(* Logix 5000 project; controller R400_500_XLS vendor 1 type 14 code 216 rev 31.11; software revision 31.01; part 15 of 32 *)
(* tags used below, declared in another part *)
   CycleModifBuffer : UDT_CYCLE;
   CycleNotEmpty : SINT;
   First_Inj_conc : BOOL;
   M : DINT[5];   // Memory Bits
   MaxTrtTempSp : REAL;
   PreWash_Select : BOOL;
   PrewashIndex : SINT;   // Index of the selected pre-wash treatment
   Rinse_Select : BOOL;
   RinseIndex : SINT;
   Second_Inj_conc : BOOL;
   Tmr : TIMER[107];
   Wash_Select : BOOL;
   WashIndex : SINT;
   WashInjectionType1 : DINT;
   CfgChem : SINT;
   CfgChem2 : SINT;
   CfgConc : REAL;
   CfgConc2 : REAL;
   CfgCondSp : REAL;
   CfgInjType : SINT;
   cfgPrewashHeated : SINT;
   cfgPrewashMin : SINT;
   cfgPrewashSec : DINT;
   CfgPrewashTempSp : REAL;
   CfgWshHeated : SINT;
   CfgWshInjRateImperial : REAL;   // Wash Injection Rate - Oz / Gal
   CfgWshInjRateMetric : REAL;   // Wash Injection Rate - mL / L
   CfgWshMin : SINT;
   CfgWshSec : SINT;
   CfgWshTempSp : REAL;
   cfgWshWport : SINT;
   ChemConcUnit : BOOL;   // 0 = mL/L; 1 = oz/gal
   Msg_TempSp : SINT;   // HMI Information Message tag
   Msg_TempSp_Ack : BOOL;
   NumInput : UDT_NUMERIC_INPUT[65];   // Numeric input
   NumInputReal : UDT_NUMERIC_INPUT_REAL[17];
   Screen_Ctrl : DINT;   // PLC Screen Request
   Selector : UDT_SELECTOR[25];   // Piloted list selector
   TempUnit : BOOL;   // Temperature Units 0= Celcius 1 = Farhenheit
   Tpb : DINT[11];
   TpbImage : DINT[11];
(* MainProgram, continued *)

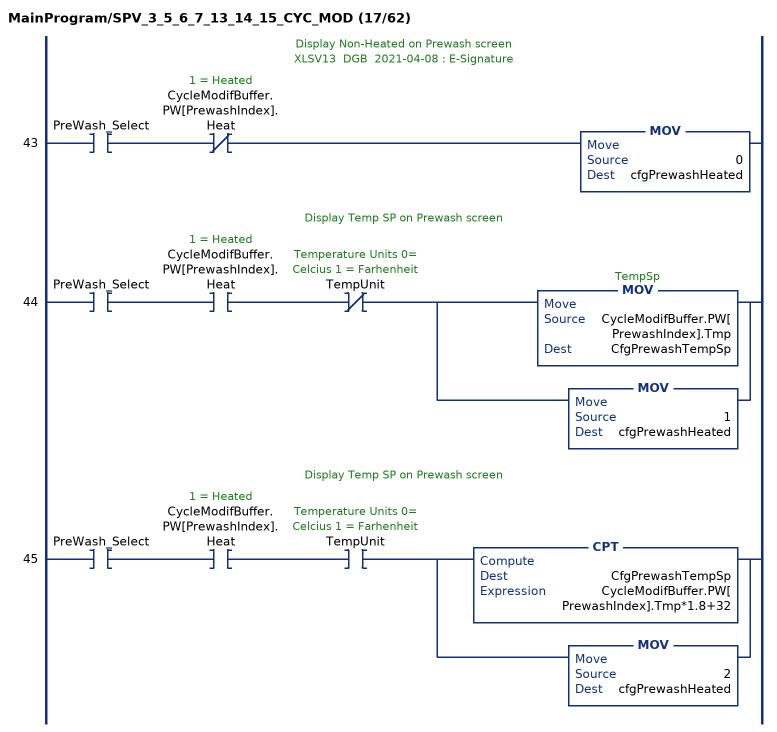
   [picture p268: MainProgram/SPV_3_5_6_7_13_14_15_CYC_MOD rungs 43-45]
   // Display Non-Heated on Prewash screen
   // XLSV13  DGB  2021-04-08 : E-Signature
   43: XIC(PreWash_Select)XIO(CycleModifBuffer.PW[PrewashIndex].Heat)MOV(0,cfgPrewashHeated);
   // Display Temp SP on Prewash screen
   44: XIC(PreWash_Select)XIC(CycleModifBuffer.PW[PrewashIndex].Heat)XIO(TempUnit)[MOV(CycleModifBuffer.PW[PrewashIndex].Tmp,CfgPrewashTempSp) ,MOV(1,cfgPrewashHeated) ];
   // Display Temp SP on Prewash screen
   45: XIC(PreWash_Select)XIC(CycleModifBuffer.PW[PrewashIndex].Heat)XIC(TempUnit)[CPT(CfgPrewashTempSp,CycleModifBuffer.PW[PrewashIndex].Tmp*1.8+32) ,MOV(2,cfgPrewashHeated) ];
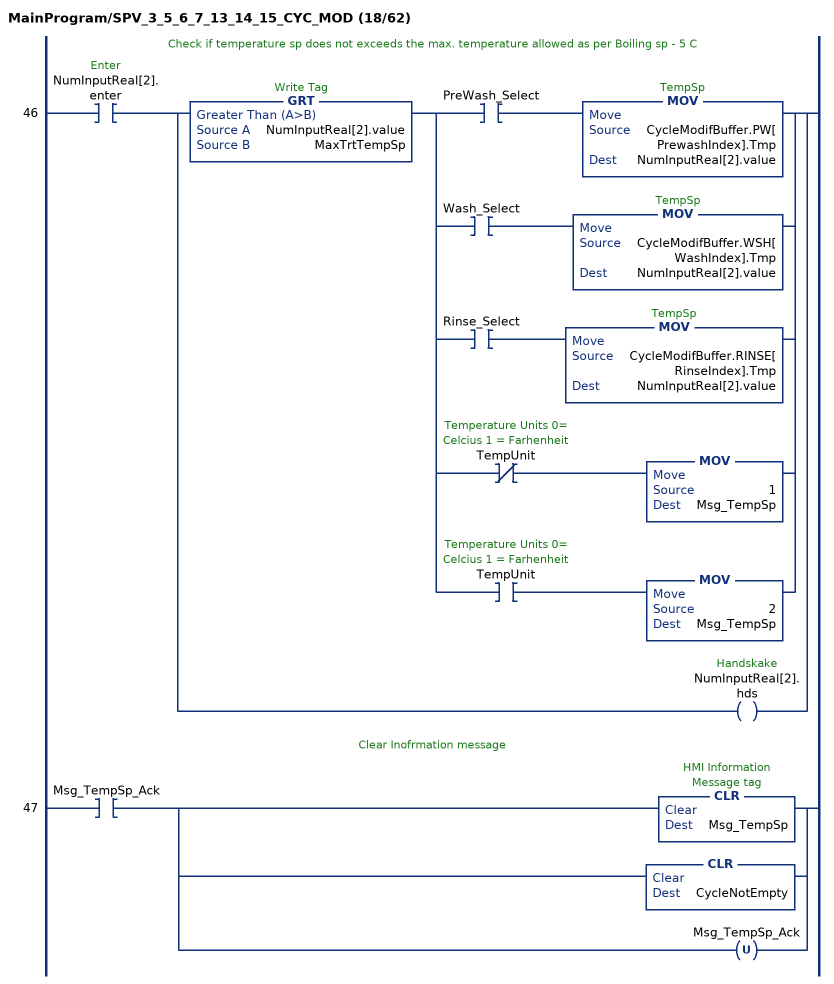
   // Check if temperature sp does not exceeds the max. temperature allowed as per Boiling sp - 5 C
   46: XIC(NumInputReal[2].enter)[GRT(NumInputReal[2].value,MaxTrtTempSp) [XIC(PreWash_Select) MOV(CycleModifBuffer.PW[PrewashIndex].Tmp,NumInputReal[2].value) ,XIC(Wash_Select) MOV(CycleModifBuffer.WSH[WashIndex].Tmp,NumInputReal[2].value) ,XIC(Rinse_Select) MOV(CycleModifBuffer.RINSE[RinseIndex].Tmp,NumInputReal[2].value) ,XIO(TempUnit) MOV(1,Msg_TempSp) ,XIC(TempUnit) MOV(2,Msg_TempSp) ] ,OTE(NumInputReal[2].hds) ];
   // Clear Inofrmation message
   47: XIC(Msg_TempSp_Ack)[CLR(Msg_TempSp) ,CLR(CycleNotEmpty) ,OTU(Msg_TempSp_Ack) ];
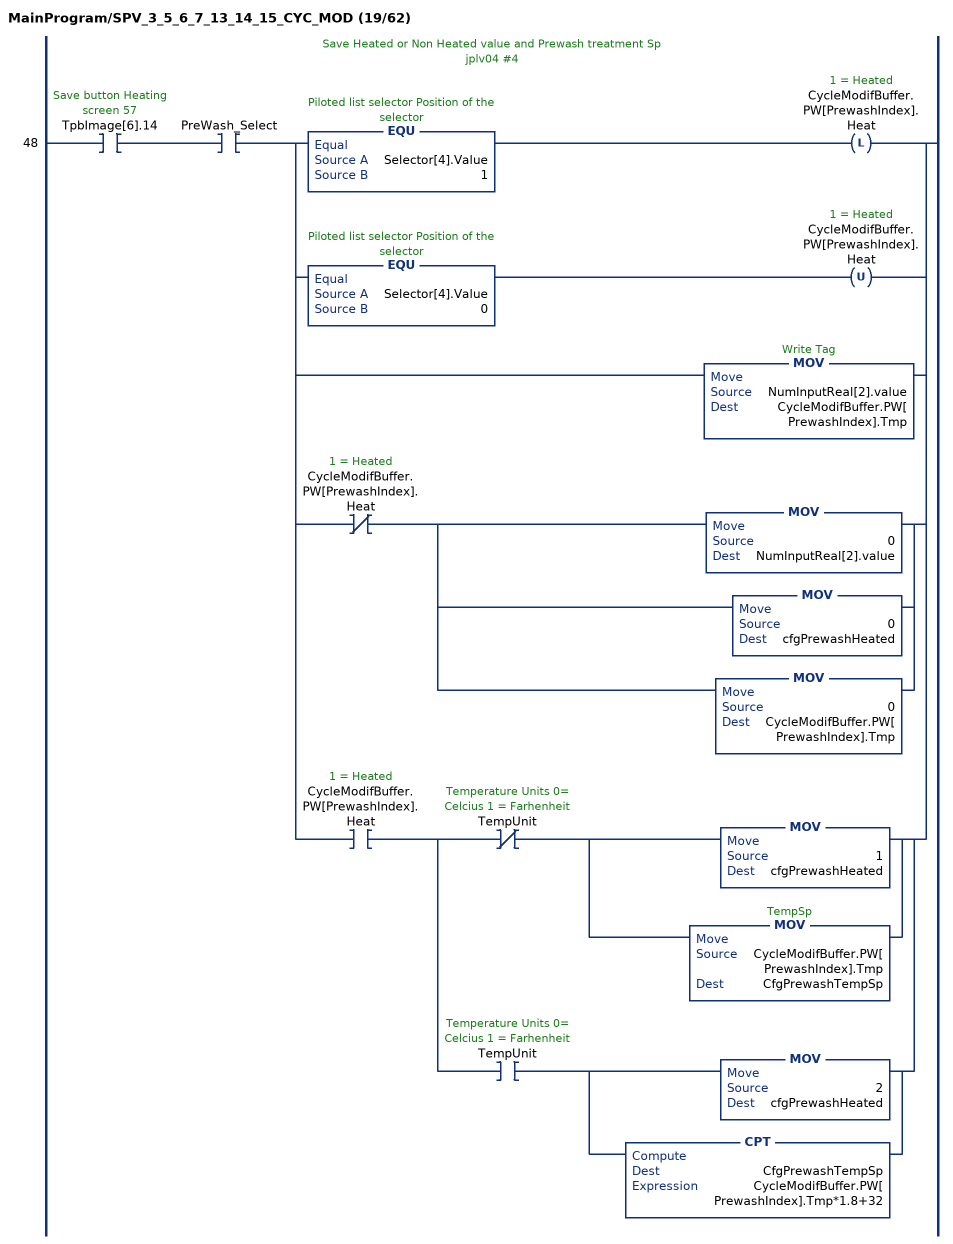
   // Save Heated or Non Heated value and Prewash treatment Sp
   // jplv04 #4
   48: XIC(TpbImage[6].14)XIC(PreWash_Select)[EQU(Selector[4].Value,1) OTL(CycleModifBuffer.PW[PrewashIndex].Heat) ,EQU(Selector[4].Value,0) OTU(CycleModifBuffer.PW[PrewashIndex].Heat) ,MOV(NumInputReal[2].value,CycleModifBuffer.PW[PrewashIndex].Tmp) ,XIO(CycleModifBuffer.PW[PrewashIndex].Heat) [MOV(0,NumInputReal[2].value) ,MOV(0,cfgPrewashHeated) ,MOV(0,CycleModifBuffer.PW[PrewashIndex].Tmp) ] ,XIC(CycleModifBuffer.PW[PrewashIndex].Heat) [XIO(TempUnit) [MOV(1,cfgPrewashHeated) ,MOV(CycleModifBuffer.PW[PrewashIndex].Tmp,CfgPrewashTempSp) ] ,XIC(TempUnit) [MOV(2,cfgPrewashHeated) ,CPT(CfgPrewashTempSp,CycleModifBuffer.PW[PrewashIndex].Tmp*1.8+32) ] ] ];
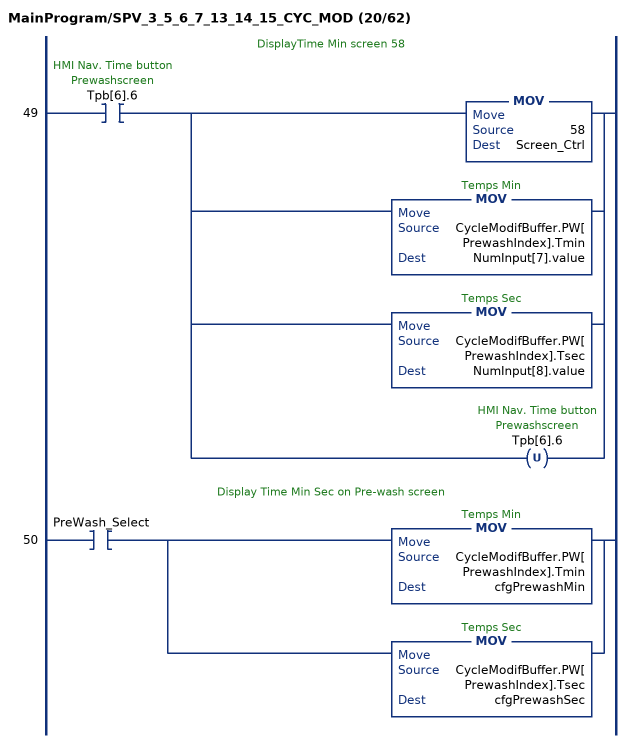
   // DisplayTime Min screen 58
   49: XIC(Tpb[6].6)[MOV(58,Screen_Ctrl) ,MOV(CycleModifBuffer.PW[PrewashIndex].Tmin,NumInput[7].value) ,MOV(CycleModifBuffer.PW[PrewashIndex].Tsec,NumInput[8].value) ,OTU(Tpb[6].6) ];
   // Display Time Min Sec on Pre-wash screen
   50: XIC(PreWash_Select)[MOV(CycleModifBuffer.PW[PrewashIndex].Tmin,cfgPrewashMin) ,MOV(CycleModifBuffer.PW[PrewashIndex].Tsec,cfgPrewashSec) ];
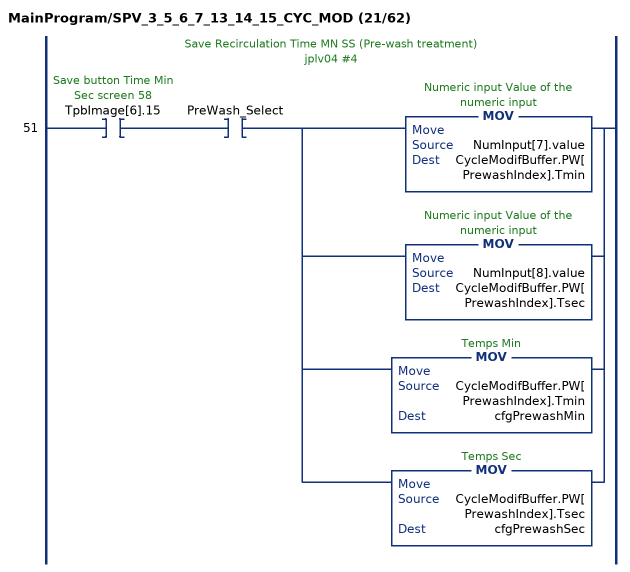
   // Save Recirculation Time MN SS (Pre-wash treatment)
   // jplv04 #4
   51: XIC(TpbImage[6].15)XIC(PreWash_Select)[MOV(NumInput[7].value,CycleModifBuffer.PW[PrewashIndex].Tmin) ,MOV(NumInput[8].value,CycleModifBuffer.PW[PrewashIndex].Tsec) ,MOV(CycleModifBuffer.PW[PrewashIndex].Tmin,cfgPrewashMin) ,MOV(CycleModifBuffer.PW[PrewashIndex].Tsec,cfgPrewashSec) ];
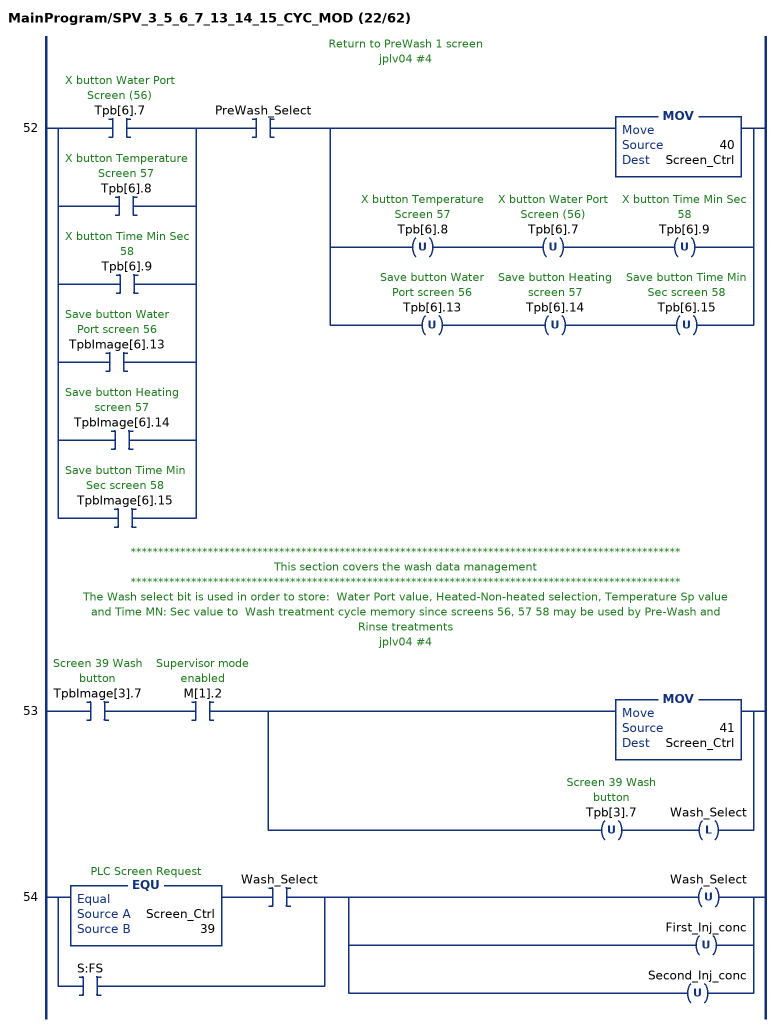
   // Return to PreWash 1 screen
   // jplv04 #4
   52: [XIC(Tpb[6].7) ,XIC(Tpb[6].8) ,XIC(Tpb[6].9) ,XIC(TpbImage[6].13) ,XIC(TpbImage[6].14) ,XIC(TpbImage[6].15) ]XIC(PreWash_Select)[MOV(40,Screen_Ctrl) ,OTU(Tpb[6].8) OTU(Tpb[6].7) OTU(Tpb[6].9) ,OTU(Tpb[6].13) OTU(Tpb[6].14) OTU(Tpb[6].15) ];
   // ****************************************************************************************************
   // This section covers the wash data management
   // ****************************************************************************************************
   // The Wash select bit is used in order to store:  Water Port value, Heated-Non-heated selection, Temperature Sp value and Time MN: Sec value to  Wash treatment cycle memory since screens 56, 57 58 may be used by Pre-Wash and Rinse treatments
   // jplv04 #4
   53: XIC(TpbImage[3].7)XIC(M[1].2)[MOV(41,Screen_Ctrl) ,OTU(Tpb[3].7) OTL(Wash_Select) ];
   54: [EQU(Screen_Ctrl,39) XIC(Wash_Select) ,XIC(S:FS) ][OTU(Wash_Select) ,OTU(First_Inj_conc) ,OTU(Second_Inj_conc) ];
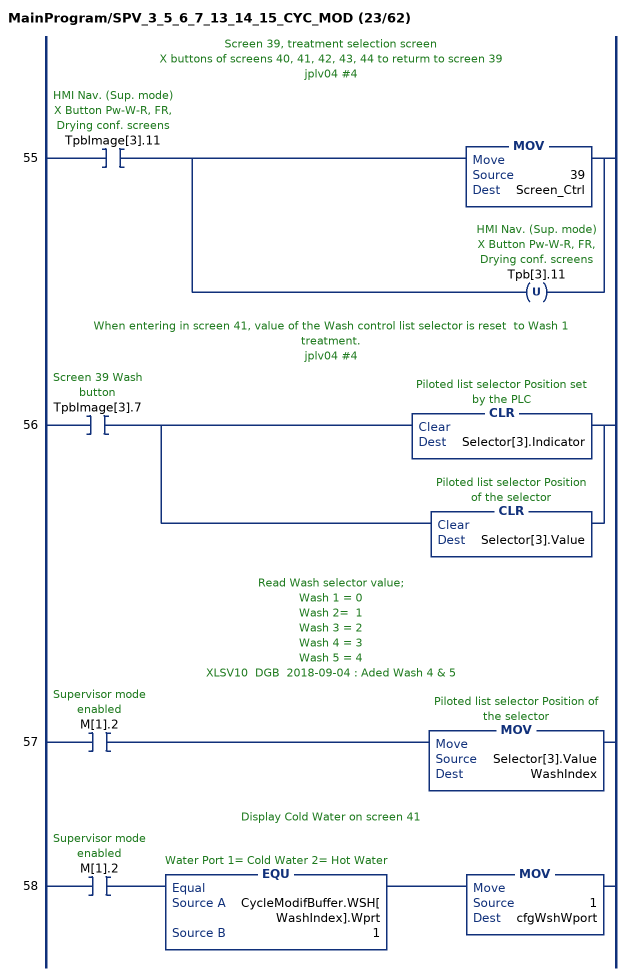
   // Screen 39, treatment selection screen
   // X buttons of screens 40, 41, 42, 43, 44 to returm to screen 39
   // jplv04 #4
   55: XIC(TpbImage[3].11)[MOV(39,Screen_Ctrl) ,OTU(Tpb[3].11) ];
   // When entering in screen 41, value of the Wash control list selector is reset  to Wash 1 treatment.
   // jplv04 #4
   56: XIC(TpbImage[3].7)[CLR(Selector[3].Indicator) ,CLR(Selector[3].Value) ];
   // Read Wash selector value;
   // Wash 1 = 0
   // Wash 2=  1
   // Wash 3 = 2
   // Wash 4 = 3
   // Wash 5 = 4
   // XLSV10  DGB  2018-09-04 : Aded Wash 4 & 5
   57: XIC(M[1].2)MOV(Selector[3].Value,WashIndex);
   // Display Cold Water on screen 41
   58: XIC(M[1].2)EQU(CycleModifBuffer.WSH[WashIndex].Wprt,1)MOV(1,cfgWshWport);
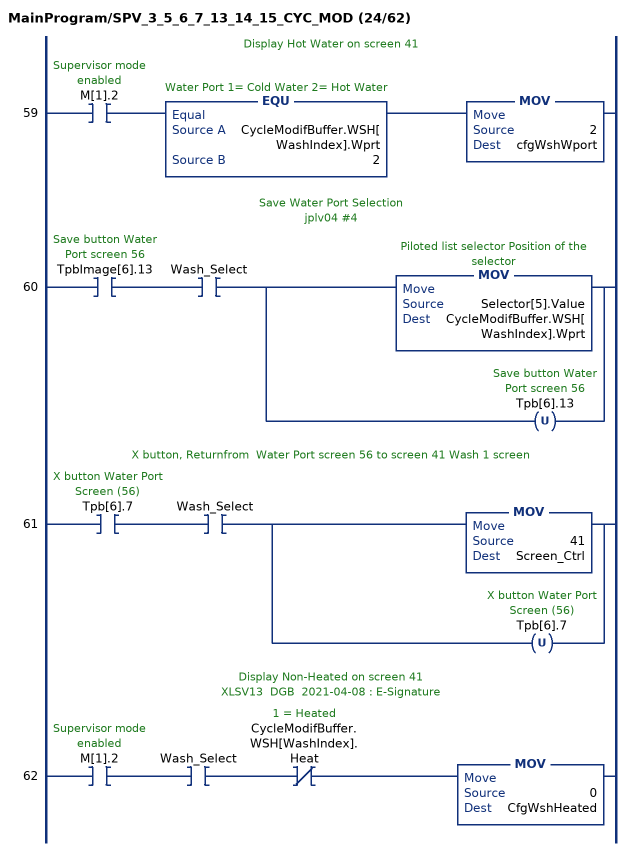
   // Display Hot Water on screen 41
   59: XIC(M[1].2)EQU(CycleModifBuffer.WSH[WashIndex].Wprt,2)MOV(2,cfgWshWport);
   // Save Water Port Selection
   // jplv04 #4
   60: XIC(TpbImage[6].13)XIC(Wash_Select)[MOV(Selector[5].Value,CycleModifBuffer.WSH[WashIndex].Wprt) ,OTU(Tpb[6].13) ];
   // X button, Returnfrom  Water Port screen 56 to screen 41 Wash 1 screen
   61: XIC(Tpb[6].7)XIC(Wash_Select)[MOV(41,Screen_Ctrl) ,OTU(Tpb[6].7) ];
   // Display Non-Heated on screen 41
   // XLSV13  DGB  2021-04-08 : E-Signature
   62: XIC(M[1].2)XIC(Wash_Select)XIO(CycleModifBuffer.WSH[WashIndex].Heat)MOV(0,CfgWshHeated);
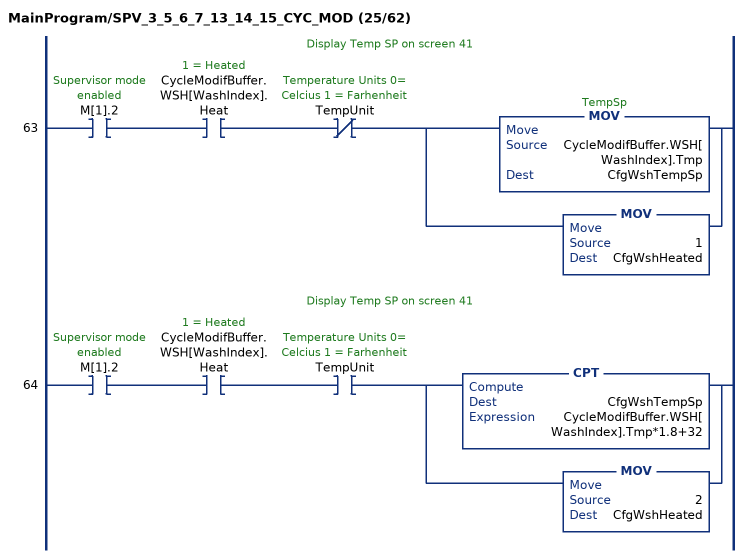
   // Display Temp SP on screen 41
   63: XIC(M[1].2)XIC(CycleModifBuffer.WSH[WashIndex].Heat)XIO(TempUnit)[MOV(CycleModifBuffer.WSH[WashIndex].Tmp,CfgWshTempSp) ,MOV(1,CfgWshHeated) ];
   // Display Temp SP on screen 41
   64: XIC(M[1].2)XIC(CycleModifBuffer.WSH[WashIndex].Heat)XIC(TempUnit)[CPT(CfgWshTempSp,CycleModifBuffer.WSH[WashIndex].Tmp*1.8+32) ,MOV(2,CfgWshHeated) ];
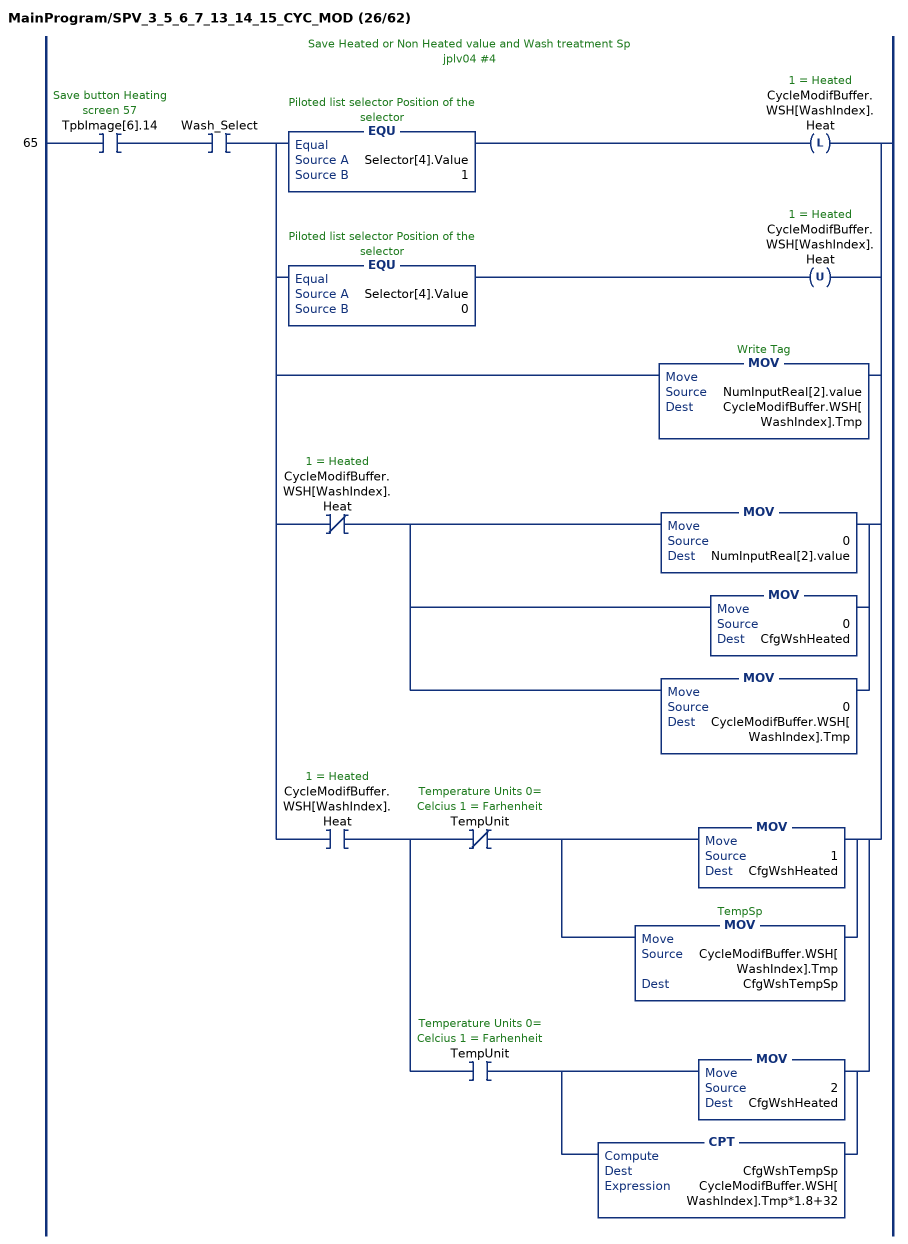
   // Save Heated or Non Heated value and Wash treatment Sp
   // jplv04 #4
   65: XIC(TpbImage[6].14)XIC(Wash_Select)[EQU(Selector[4].Value,1) OTL(CycleModifBuffer.WSH[WashIndex].Heat) ,EQU(Selector[4].Value,0) OTU(CycleModifBuffer.WSH[WashIndex].Heat) ,MOV(NumInputReal[2].value,CycleModifBuffer.WSH[WashIndex].Tmp) ,XIO(CycleModifBuffer.WSH[WashIndex].Heat) [MOV(0,NumInputReal[2].value) ,MOV(0,CfgWshHeated) ,MOV(0,CycleModifBuffer.WSH[WashIndex].Tmp) ] ,XIC(CycleModifBuffer.WSH[WashIndex].Heat) [XIO(TempUnit) [MOV(1,CfgWshHeated) ,MOV(CycleModifBuffer.WSH[WashIndex].Tmp,CfgWshTempSp) ] ,XIC(TempUnit) [MOV(2,CfgWshHeated) ,CPT(CfgWshTempSp,CycleModifBuffer.WSH[WashIndex].Tmp*1.8+32) ] ] ];
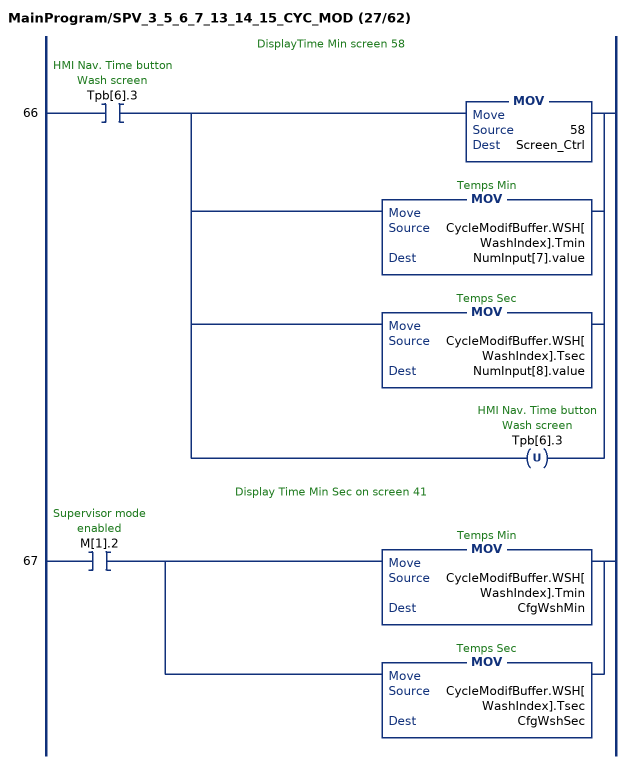
   // DisplayTime Min screen 58
   66: XIC(Tpb[6].3)[MOV(58,Screen_Ctrl) ,MOV(CycleModifBuffer.WSH[WashIndex].Tmin,NumInput[7].value) ,MOV(CycleModifBuffer.WSH[WashIndex].Tsec,NumInput[8].value) ,OTU(Tpb[6].3) ];
   // Display Time Min Sec on screen 41
   67: XIC(M[1].2)[MOV(CycleModifBuffer.WSH[WashIndex].Tmin,CfgWshMin) ,MOV(CycleModifBuffer.WSH[WashIndex].Tsec,CfgWshSec) ];
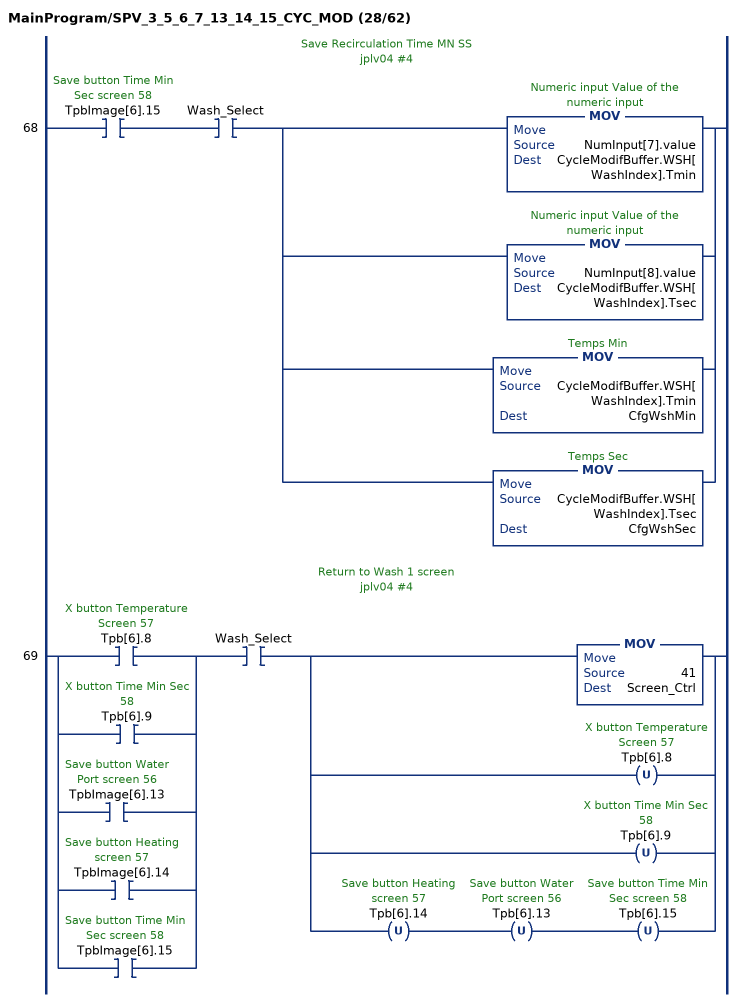
   // Save Recirculation Time MN SS
   // jplv04 #4
   68: XIC(TpbImage[6].15)XIC(Wash_Select)[MOV(NumInput[7].value,CycleModifBuffer.WSH[WashIndex].Tmin) ,MOV(NumInput[8].value,CycleModifBuffer.WSH[WashIndex].Tsec) ,MOV(CycleModifBuffer.WSH[WashIndex].Tmin,CfgWshMin) ,MOV(CycleModifBuffer.WSH[WashIndex].Tsec,CfgWshSec) ];
   // Return to Wash 1 screen
   // jplv04 #4
   69: [XIC(Tpb[6].8) ,XIC(Tpb[6].9) ,XIC(TpbImage[6].13) ,XIC(TpbImage[6].14) ,XIC(TpbImage[6].15) ]XIC(Wash_Select)[MOV(41,Screen_Ctrl) ,OTU(Tpb[6].8) ,OTU(Tpb[6].9) ,OTU(Tpb[6].14) OTU(Tpb[6].13) OTU(Tpb[6].15) ];
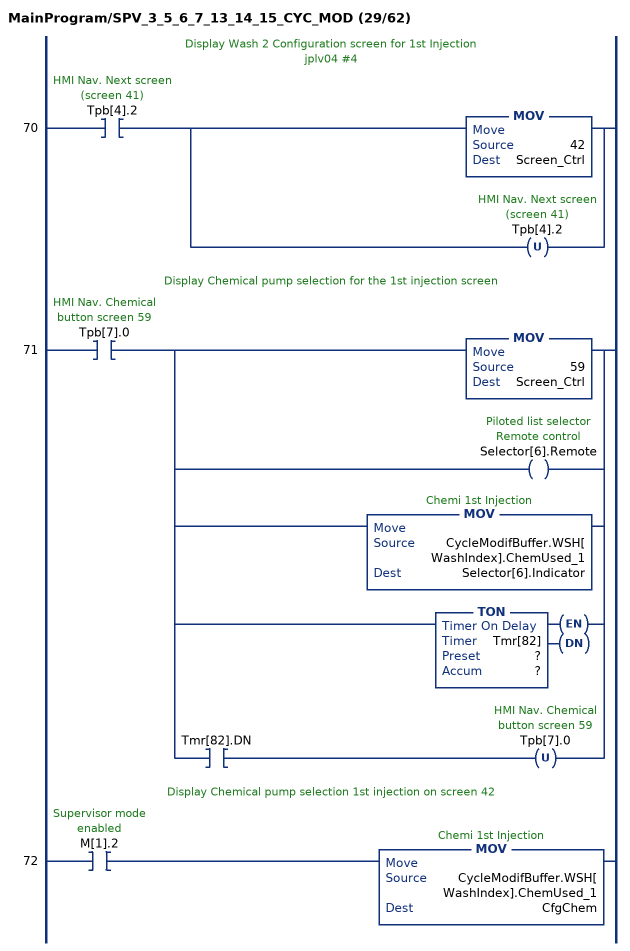
   // Display Wash 2 Configuration screen for 1st Injection
   // jplv04 #4
   70: XIC(Tpb[4].2)[MOV(42,Screen_Ctrl) ,OTU(Tpb[4].2) ];
   // Display Chemical pump selection for the 1st injection screen
   71: XIC(Tpb[7].0)[MOV(59,Screen_Ctrl) ,OTE(Selector[6].Remote) ,MOV(CycleModifBuffer.WSH[WashIndex].ChemUsed_1,Selector[6].Indicator) ,TON(Tmr[82],?,?) ,XIC(Tmr[82].DN) OTU(Tpb[7].0) ];
   // Display Chemical pump selection 1st injection on screen 42
   72: XIC(M[1].2)MOV(CycleModifBuffer.WSH[WashIndex].ChemUsed_1,CfgChem);
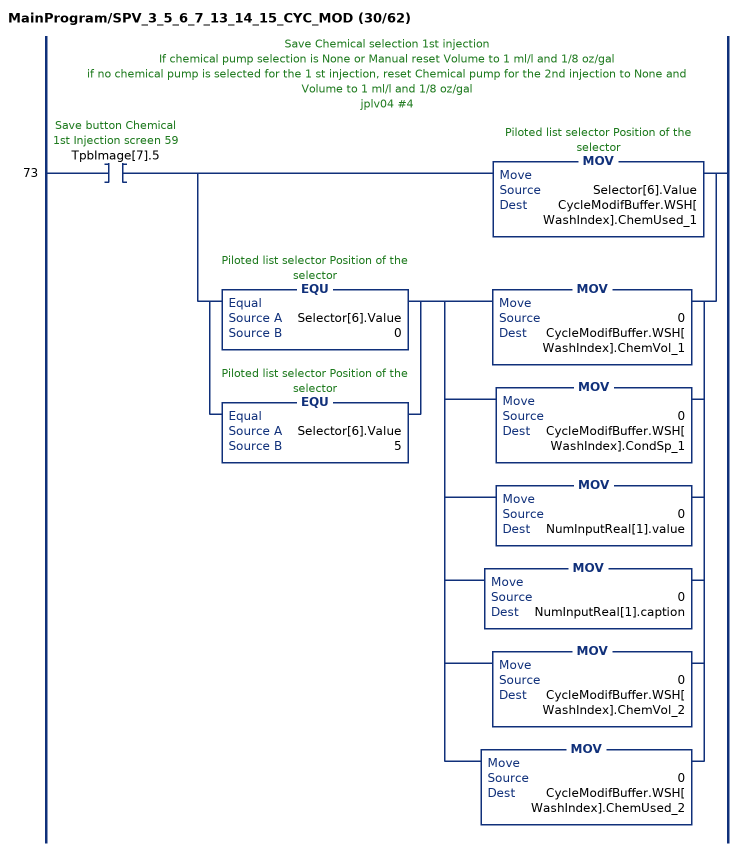
   // Save Chemical selection 1st injection
   // If chemical pump selection is None or Manual reset Volume to 1 ml/l and 1/8 oz/gal
   // if no chemical pump is selected for the 1 st injection, reset Chemical pump for the 2nd injection to None and Volume to 1 ml/l and 1/8 oz/gal
   // jplv04 #4
   73: XIC(TpbImage[7].5)[MOV(Selector[6].Value,CycleModifBuffer.WSH[WashIndex].ChemUsed_1) ,[EQU(Selector[6].Value,0) ,EQU(Selector[6].Value,5) ] [MOV(0,CycleModifBuffer.WSH[WashIndex].ChemVol_1) ,MOV(0,CycleModifBuffer.WSH[WashIndex].CondSp_1) ,MOV(0,NumInputReal[1].value) ,MOV(0,NumInputReal[1].caption) ,MOV(0,CycleModifBuffer.WSH[WashIndex].ChemVol_2) ,MOV(0,CycleModifBuffer.WSH[WashIndex].ChemUsed_2) ] ];
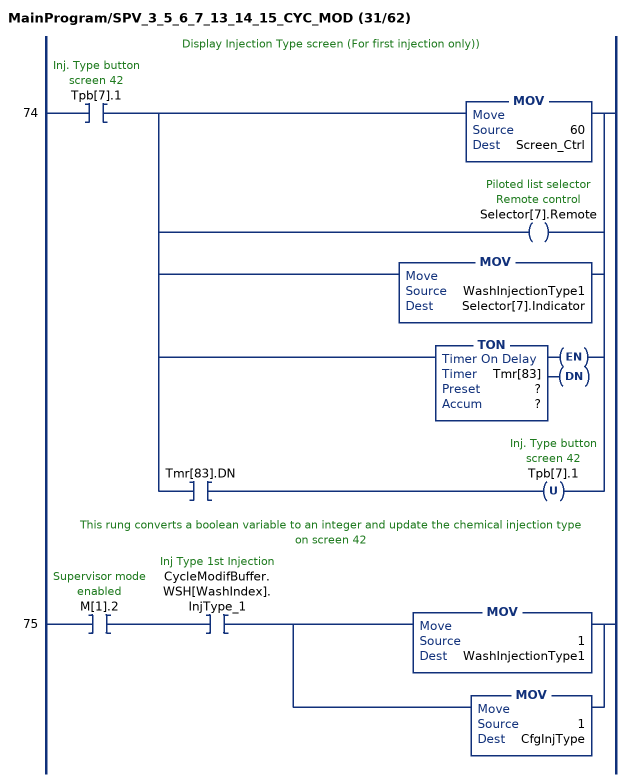
   // Display Injection Type screen (For first injection only))
   74: XIC(Tpb[7].1)[MOV(60,Screen_Ctrl) ,OTE(Selector[7].Remote) ,MOV(WashInjectionType1,Selector[7].Indicator) ,TON(Tmr[83],?,?) ,XIC(Tmr[83].DN) OTU(Tpb[7].1) ];
   // This rung converts a boolean variable to an integer and update the chemical injection type on screen 42
   75: XIC(M[1].2)XIC(CycleModifBuffer.WSH[WashIndex].InjType_1)[MOV(1,WashInjectionType1) ,MOV(1,CfgInjType) ];
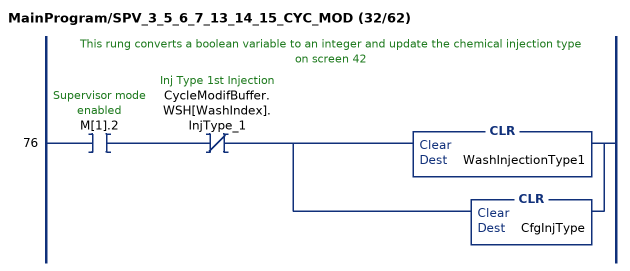
   // This rung converts a boolean variable to an integer and update the chemical injection type on screen 42
   76: XIC(M[1].2)XIO(CycleModifBuffer.WSH[WashIndex].InjType_1)[CLR(WashInjectionType1) ,CLR(CfgInjType) ];
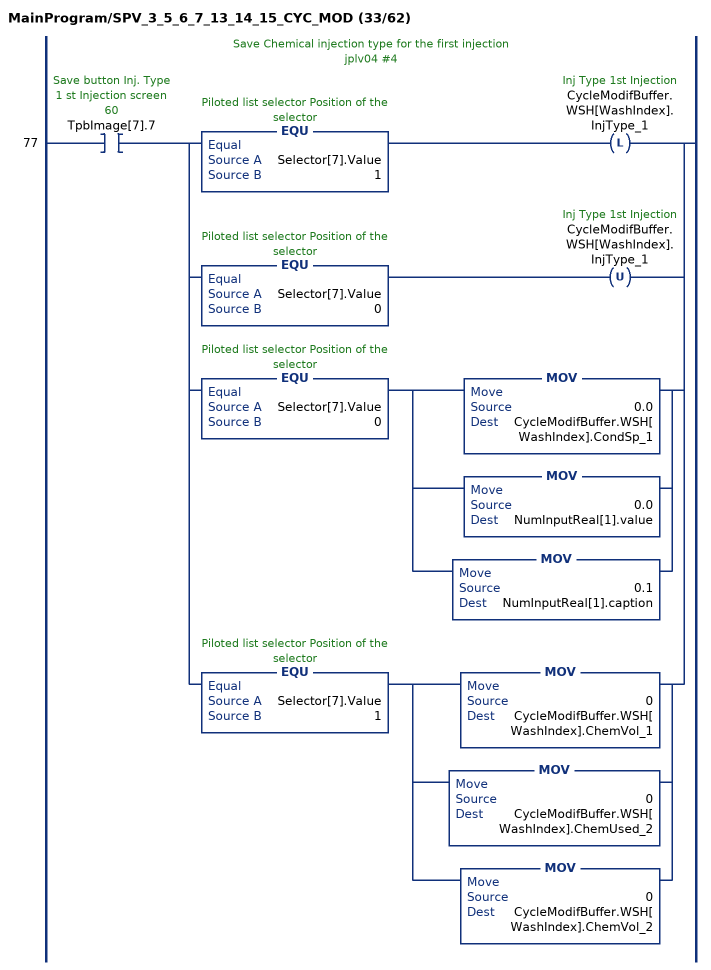
   // Save Chemical injection type for the first injection
   // jplv04 #4
   77: XIC(TpbImage[7].7)[EQU(Selector[7].Value,1) OTL(CycleModifBuffer.WSH[WashIndex].InjType_1) ,EQU(Selector[7].Value,0) OTU(CycleModifBuffer.WSH[WashIndex].InjType_1) ,EQU(Selector[7].Value,0) [MOV(0.0,CycleModifBuffer.WSH[WashIndex].CondSp_1) ,MOV(0.0,NumInputReal[1].value) ,MOV(0.1,NumInputReal[1].caption) ] ,EQU(Selector[7].Value,1) [MOV(0,CycleModifBuffer.WSH[WashIndex].ChemVol_1) ,MOV(0,CycleModifBuffer.WSH[WashIndex].ChemUsed_2) ,MOV(0,CycleModifBuffer.WSH[WashIndex].ChemVol_2) ] ];
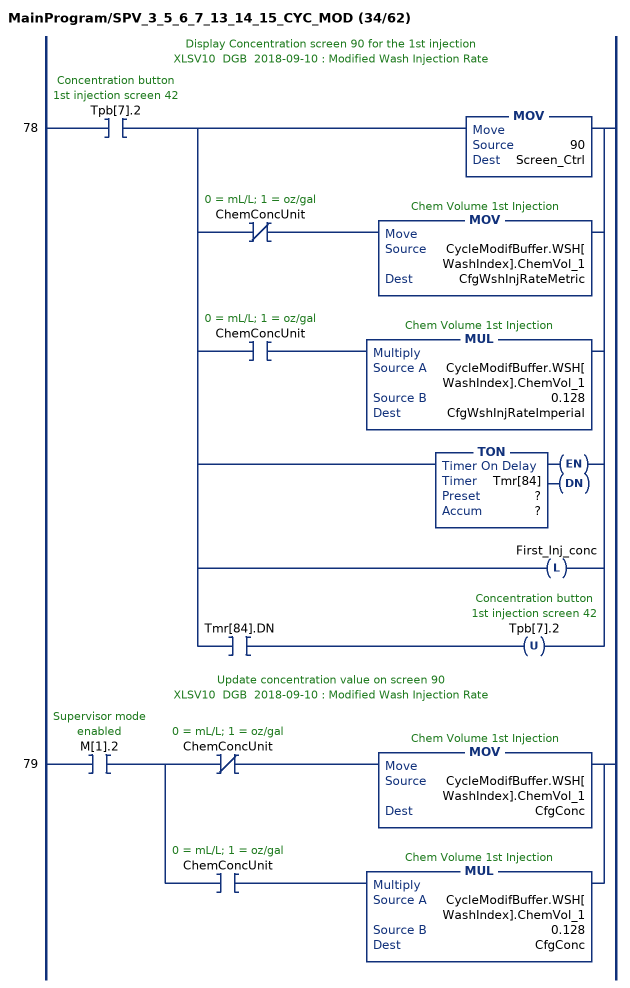
   // Display Concentration screen 90 for the 1st injection
   // XLSV10  DGB  2018-09-10 : Modified Wash Injection Rate
   78: XIC(Tpb[7].2)[MOV(90,Screen_Ctrl) ,XIO(ChemConcUnit) MOV(CycleModifBuffer.WSH[WashIndex].ChemVol_1,CfgWshInjRateMetric) ,XIC(ChemConcUnit) MUL(CycleModifBuffer.WSH[WashIndex].ChemVol_1,0.128,CfgWshInjRateImperial) ,TON(Tmr[84],?,?) ,OTL(First_Inj_conc) ,XIC(Tmr[84].DN) OTU(Tpb[7].2) ];
   // Update concentration value on screen 90
   // XLSV10  DGB  2018-09-10 : Modified Wash Injection Rate
   79: XIC(M[1].2)[XIO(ChemConcUnit) MOV(CycleModifBuffer.WSH[WashIndex].ChemVol_1,CfgConc) ,XIC(ChemConcUnit) MUL(CycleModifBuffer.WSH[WashIndex].ChemVol_1,0.128,CfgConc) ];
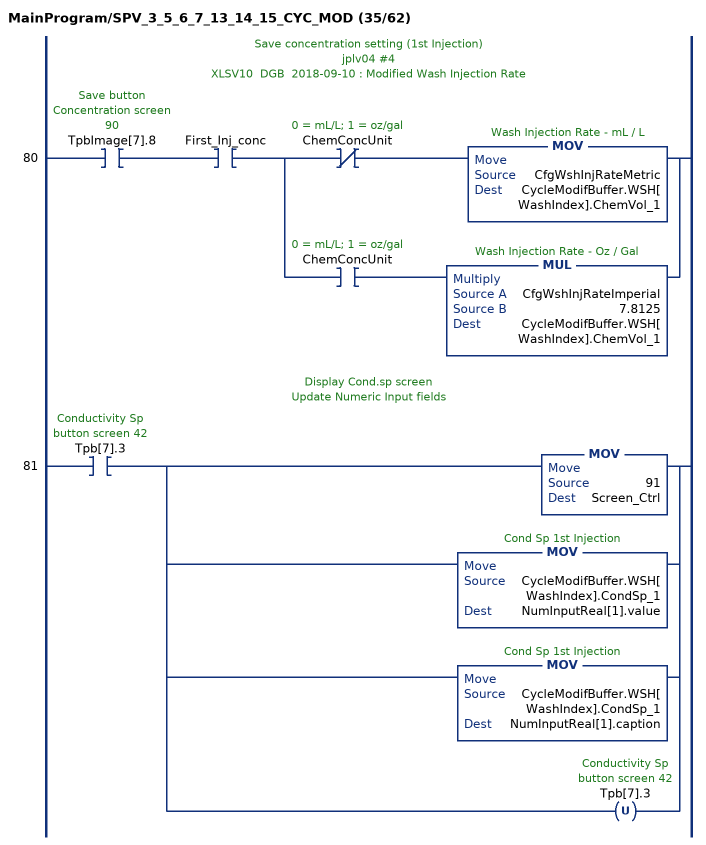
   // Save concentration setting (1st Injection)
   // jplv04 #4
   // XLSV10  DGB  2018-09-10 : Modified Wash Injection Rate
   80: XIC(TpbImage[7].8)XIC(First_Inj_conc)[XIO(ChemConcUnit) MOV(CfgWshInjRateMetric,CycleModifBuffer.WSH[WashIndex].ChemVol_1) ,XIC(ChemConcUnit) MUL(CfgWshInjRateImperial,7.8125,CycleModifBuffer.WSH[WashIndex].ChemVol_1) ];
   // Display Cond.sp screen
   // Update Numeric Input fields
   81: XIC(Tpb[7].3)[MOV(91,Screen_Ctrl) ,MOV(CycleModifBuffer.WSH[WashIndex].CondSp_1,NumInputReal[1].value) ,MOV(CycleModifBuffer.WSH[WashIndex].CondSp_1,NumInputReal[1].caption) ,OTU(Tpb[7].3) ];
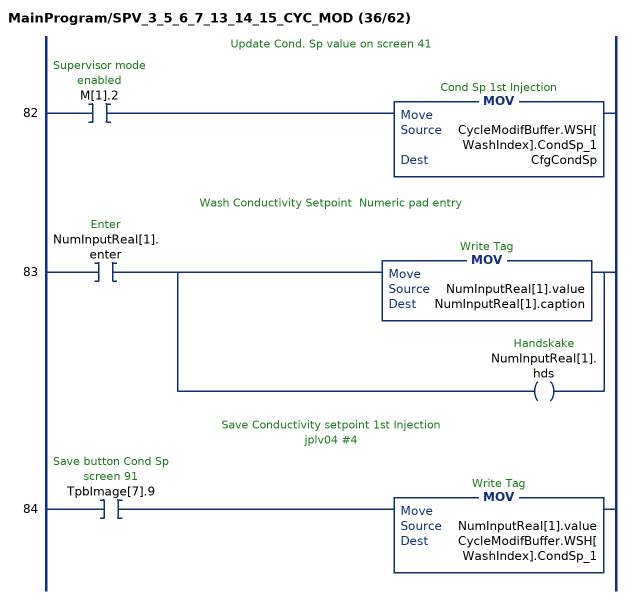
   // Update Cond. Sp value on screen 41
   82: XIC(M[1].2)MOV(CycleModifBuffer.WSH[WashIndex].CondSp_1,CfgCondSp);
   // Wash Conductivity Setpoint  Numeric pad entry
   83: XIC(NumInputReal[1].enter)[MOV(NumInputReal[1].value,NumInputReal[1].caption) ,OTE(NumInputReal[1].hds) ];
   // Save Conductivity setpoint 1st Injection
   // jplv04 #4
   84: XIC(TpbImage[7].9)MOV(NumInputReal[1].value,CycleModifBuffer.WSH[WashIndex].CondSp_1);
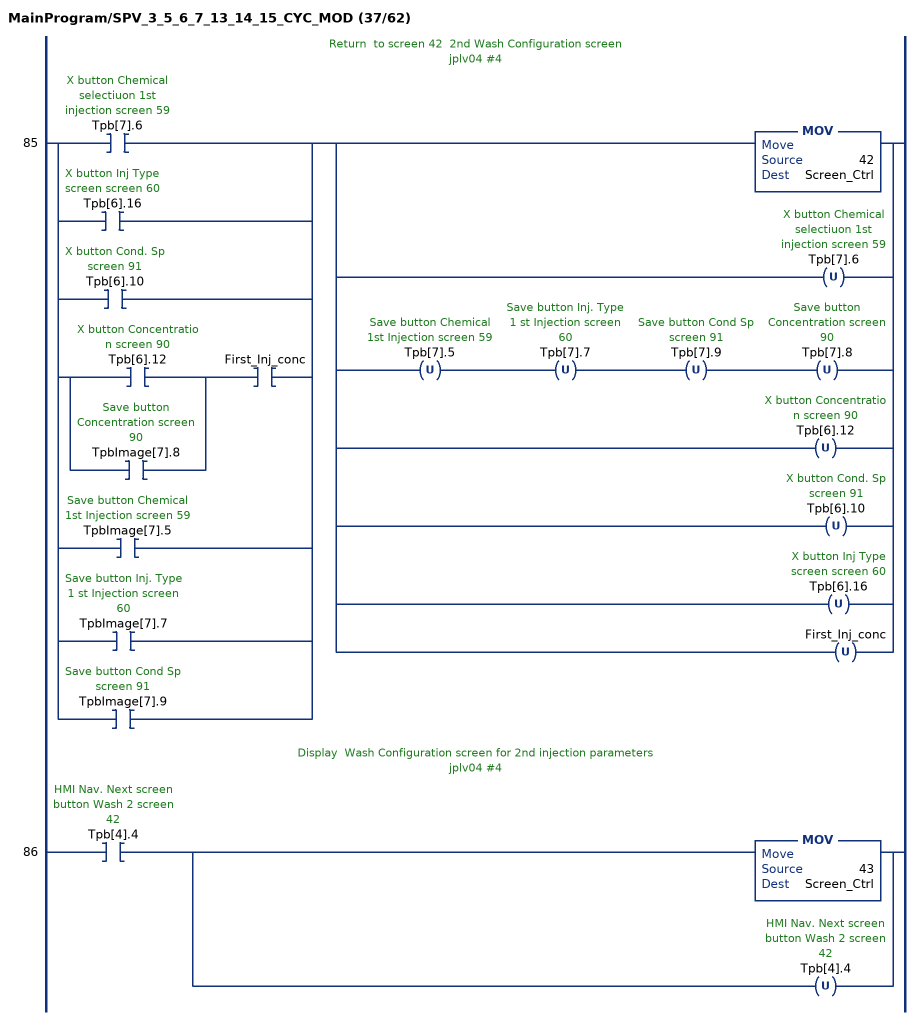
   // Return  to screen 42  2nd Wash Configuration screen
   // jplv04 #4
   85: [XIC(Tpb[7].6) ,XIC(Tpb[6].16) ,XIC(Tpb[6].10) ,[XIC(Tpb[6].12) ,XIC(TpbImage[7].8) ] XIC(First_Inj_conc) ,XIC(TpbImage[7].5) ,XIC(TpbImage[7].7) ,XIC(TpbImage[7].9) ][MOV(42,Screen_Ctrl) ,OTU(Tpb[7].6) ,OTU(Tpb[7].5) OTU(Tpb[7].7) OTU(Tpb[7].9) OTU(Tpb[7].8) ,OTU(Tpb[6].12) ,OTU(Tpb[6].10) ,OTU(Tpb[6].16) ,OTU(First_Inj_conc) ];
   // Display  Wash Configuration screen for 2nd injection parameters
   // jplv04 #4
   86: XIC(Tpb[4].4)[MOV(43,Screen_Ctrl) ,OTU(Tpb[4].4) ];
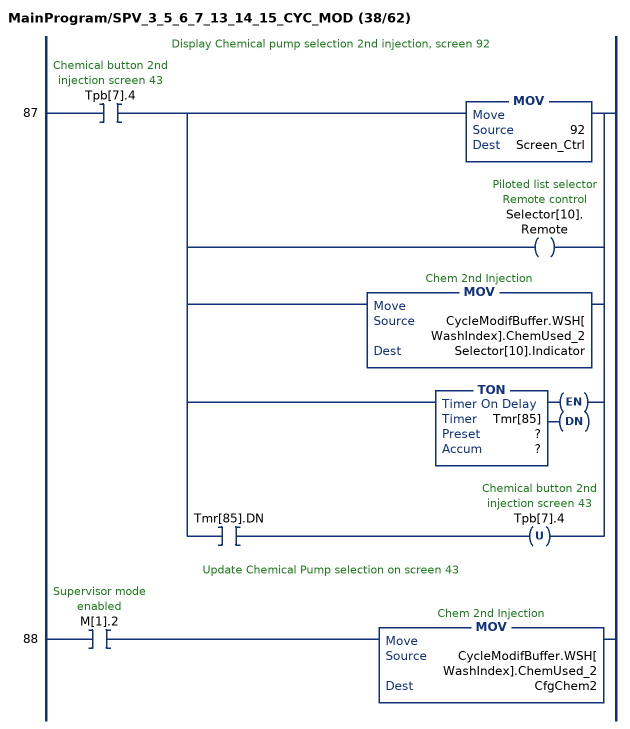
   // Display Chemical pump selection 2nd injection, screen 92
   87: XIC(Tpb[7].4)[MOV(92,Screen_Ctrl) ,OTE(Selector[10].Remote) ,MOV(CycleModifBuffer.WSH[WashIndex].ChemUsed_2,Selector[10].Indicator) ,TON(Tmr[85],?,?) ,XIC(Tmr[85].DN) OTU(Tpb[7].4) ];
   // Update Chemical Pump selection on screen 43
   88: XIC(M[1].2)MOV(CycleModifBuffer.WSH[WashIndex].ChemUsed_2,CfgChem2);
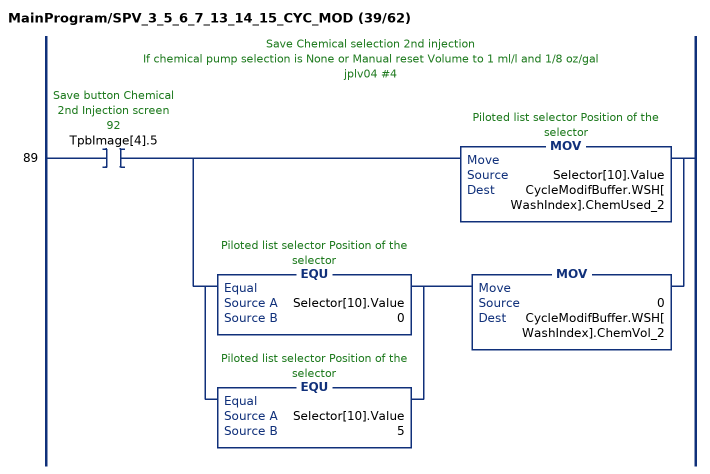
   // Save Chemical selection 2nd injection
   // If chemical pump selection is None or Manual reset Volume to 1 ml/l and 1/8 oz/gal
   // jplv04 #4
   89: XIC(TpbImage[4].5)[MOV(Selector[10].Value,CycleModifBuffer.WSH[WashIndex].ChemUsed_2) ,[EQU(Selector[10].Value,0) ,EQU(Selector[10].Value,5) ] MOV(0,CycleModifBuffer.WSH[WashIndex].ChemVol_2) ];
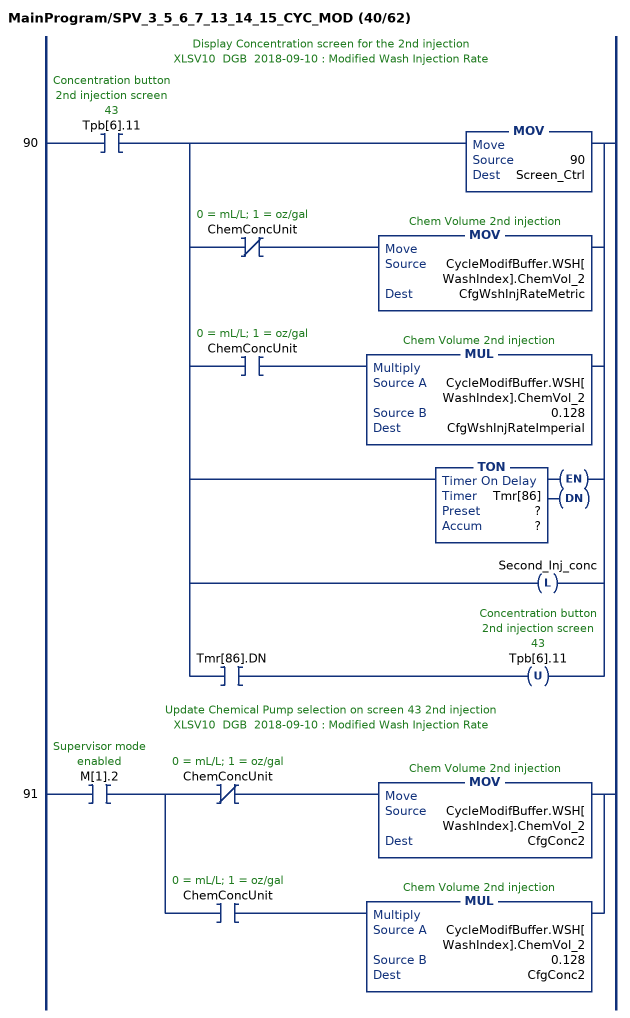
   // Display Concentration screen for the 2nd injection
   // XLSV10  DGB  2018-09-10 : Modified Wash Injection Rate
   90: XIC(Tpb[6].11)[MOV(90,Screen_Ctrl) ,XIO(ChemConcUnit) MOV(CycleModifBuffer.WSH[WashIndex].ChemVol_2,CfgWshInjRateMetric) ,XIC(ChemConcUnit) MUL(CycleModifBuffer.WSH[WashIndex].ChemVol_2,0.128,CfgWshInjRateImperial) ,TON(Tmr[86],?,?) ,OTL(Second_Inj_conc) ,XIC(Tmr[86].DN) OTU(Tpb[6].11) ];
   // Update Chemical Pump selection on screen 43 2nd injection
   // XLSV10  DGB  2018-09-10 : Modified Wash Injection Rate
   91: XIC(M[1].2)[XIO(ChemConcUnit) MOV(CycleModifBuffer.WSH[WashIndex].ChemVol_2,CfgConc2) ,XIC(ChemConcUnit) MUL(CycleModifBuffer.WSH[WashIndex].ChemVol_2,0.128,CfgConc2) ];
